(* IEC 61131-3 sources: courses/root/cat/cat-hw-boards/safety-plc/proj-safety-plc-emergency-stop-integration/structured-text, 4 files *)

(* ---- SafetyTypes.st ---- *)
TYPE E_SafetyState :
(
    STATE_SAFE := 0,               (* Безпечний робочий стан, силові виходи увімкнені *)
    STATE_ESTOP_ACTIVE := 1,        (* Натиснуто кнопку аварійної зупинки E-Stop (канали розімкнені) *)
    STATE_WAITING_FOR_RESET := 2,    (* Входи відновлено, очікується ручне підтвердження (Reset) *)
    STATE_DISCREPANCY_FAULT := 3,   (* Апаратна помилка: перевищено час розбіжності між каналами *)
    STATE_EDM_FAULT := 4            (* Апаратна помилка: несправність контактора або приварювання контактів *)
);
END_TYPE

TYPE E_EStopFault :
(
    ESTOP_FAULT_NONE := 0,                 (* Помилки відсутні *)
    ESTOP_FAULT_DISCREPANCY_TIMEOUT := 1,   (* Перевищення часу розбіжності спрацьовування каналів *)
    ESTOP_FAULT_EDM := 2,                   (* Несправність ланцюга зворотного зв'язку EDM *)
    ESTOP_FAULT_INVALID_RESET := 3          (* Некоректна послідовність скидання *)
);
END_TYPE

TYPE E_EdmFaultState :
(
    EDM_FAULT_NONE := 0,                (* Ланцюг зворотного зв'язку справний *)
    EDM_FAULT_CONTACT_WELDED := 1,      (* Приварювання контактів (NC не замкнувся при вимкненні) *)
    EDM_FAULT_CONTACT_STUCK_OPEN := 2,  (* Заклинювання реле (NC не розімкнувся при увімкненні) *)
    EDM_FAULT_TIMEOUT := 3              (* Таймаут підтвердження стану контакторів *)
);
END_TYPE

TYPE ST_EdmConfig :
STRUCT
    tFeedbackTimeout : TIME := T#250ms; (* Максимальний час очікування відповіді зворотного зв'язку *)
END_STRUCT
END_TYPE

TYPE ST_EStopConfig :
STRUCT
    tDiscrepancyTime : TIME := T#100ms; (* Допустима часова розбіжність між каналами E-Stop *)
    stEdmConfig      : ST_EdmConfig;    (* Конфігурація моніторингу зворотного зв'язку *)
END_STRUCT
END_TYPE

(* ---- FB_EDM_Monitor.st ---- *)
(*
    Функціональний блок: FB_EDM_Monitor
    Опис: Здійснює моніторинг зворотного зв'язку (External Device Monitoring) силових контакторів
          через їхні розмикальні (NC) допоміжні контакти. Забезпечує виявлення заклинювання
          або приварювання контактів за допомогою таймера контролю допустимої затримки перемикання.
*)
FUNCTION_BLOCK FB_EDM_Monitor
VAR_INPUT
    bControlOutput : BOOL;          (* Сигнал керування силових виходів (TRUE = увімкнено, FALSE = вимкнено) *)
    bFeedbackNC    : BOOL;          (* Сигнал з розмикальних (NC) допоміжних контактів контактора *)
    bReset         : BOOL;          (* Сигнал скидання помилки EDM *)
    stConfig       : ST_EdmConfig;  (* Конфігурація таймаутів моніторингу *)
END_VAR
VAR_OUTPUT
    bEdmOk         : BOOL := FALSE; (* Прапор норми: TRUE = ланцюг зворотного зв'язку у належному стані *)
    bError         : BOOL := FALSE; (* Прапор фіксації апаратної помилки контакторів *)
    eFaultState    : E_EdmFaultState := E_EdmFaultState.EDM_FAULT_NONE; (* Тип діагностованої помилки *)
END_VAR
VAR
    timerDelay     : TON;           (* Таймер затримки перемикання контактів *)
    bMismatch      : BOOL;          (* Прапор розбіжності між командою та зворотним зв'язком *)
END_VAR

(*
    Логіка моніторингу:
    У стабільному стані стан NC-контакту має бути протилежним команді керування:
    - Якщо bControlOutput = FALSE (контактор знеструмлено), NC-контакт має замкнутися (bFeedbackNC = TRUE).
    - Якщо bControlOutput = TRUE (контактор під напругою), NC-контакт має розімкнутися (bFeedbackNC = FALSE).
    Якщо bControlOutput = bFeedbackNC, виникає невідповідність (bMismatch = TRUE).
*)
bMismatch := (bControlOutput = bFeedbackNC);

(* Запуск таймера перевірки затримки спрацьовування *)
timerDelay(IN := bMismatch AND NOT bError, PT := stConfig.tFeedbackTimeout);

(* Фіксація помилки у разі перевищення таймауту *)
IF timerDelay.Q THEN
    bError := TRUE;
    IF NOT bControlOutput AND NOT bFeedbackNC THEN
        (* Вихід вимкнено, але NC-контакт не замкнувся -> приварювання силових контактів *)
        eFaultState := E_EdmFaultState.EDM_FAULT_CONTACT_WELDED;
    ELSIF bControlOutput AND bFeedbackNC THEN
        (* Вихід увімкнено, але NC-контакт не розімкнувся -> заклинювання у розімкненому стані *)
        eFaultState := E_EdmFaultState.EDM_FAULT_CONTACT_STUCK_OPEN;
    ELSE
        eFaultState := E_EdmFaultState.EDM_FAULT_TIMEOUT;
    END_IF;
END_IF;

(* Обробка процедури скидання помилки *)
IF bReset THEN
    (* Скидання дозволено лише якщо команду вимкнено і NC-контакт дійсно відновлено (замкнено) *)
    IF NOT bControlOutput AND bFeedbackNC THEN
        bError := FALSE;
        eFaultState := E_EdmFaultState.EDM_FAULT_NONE;
    END_IF;
END_IF;

(* Формування підсумкового прапорця стану EDM *)
bEdmOk := NOT bError AND NOT timerDelay.Q AND NOT bMismatch;

END_FUNCTION_BLOCK

(* ---- FB_EStop.st ---- *)
(*
    Функціональний блок: FB_EStop
    Опис: Реалізує функціонал безпеки двоканального аварійного зупину (E-Stop) з перевіркою
          часової розбіжності входів (Discrepancy Time), інтегрованим моніторингом зворотного
          зв'язку силових реле (EDM) та детермінованим автоматом станів.
*)
FUNCTION_BLOCK FB_EStop
VAR_INPUT
    bChannel1      : BOOL;          (* Перший канал кнопки E-Stop (F-DI 1, NC) *)
    bChannel2      : BOOL;          (* Другий канал кнопки E-Stop (F-DI 2, NC) *)
    bFeedbackNC    : BOOL;          (* Зворотний зв'язок NC-контактів силових реле *)
    bReset         : BOOL;          (* Сигнал кнопки ручного підтвердження/скидання (Reset) *)
    stConfig       : ST_EStopConfig;(* Параметри затримок та конфігурація EDM *)
END_VAR
VAR_OUTPUT
    bSafetyOutput  : BOOL := FALSE; (* Вихід дозволу роботи силових ланцюгів (F-DO) *)
    bReadyForReset : BOOL := FALSE; (* Сигнал індикації готовності до скидання (очікування Reset) *)
    bError         : BOOL := FALSE; (* Прапор виявлення апаратної помилки *)
    eState         : E_SafetyState := E_SafetyState.STATE_ESTOP_ACTIVE; (* Поточний стан безпеки *)
    eFault         : E_EStopFault  := E_EStopFault.ESTOP_FAULT_NONE;    (* Поточна фіксована помилка *)
END_VAR
VAR
    fbEdm          : FB_EDM_Monitor;(* Екземпляр блоку моніторингу контакторів *)
    timerDiscrepancy: TON;          (* Таймер контролю часової розбіжності входів *)
    rTrigReset     : R_TRIG;        (* Визначник наростаючого фронту для сигналу Reset *)
END_VAR

(* Виявлення фронту сигналу скидання (захист від постійно затиснутої кнопки Reset) *)
rTrigReset(CLK := bReset);

(* Виклик підсистеми EDM моніторингу *)
fbEdm(
    bControlOutput := bSafetyOutput,
    bFeedbackNC    := bFeedbackNC,
    bReset         := bReset,
    stConfig       := stConfig.stEdmConfig
);

(* Таймер контролю часової розбіжності між двома каналами кнопки аварійної зупинки *)
timerDiscrepancy(
    IN := (bChannel1 <> bChannel2) AND (eState <> E_SafetyState.STATE_DISCREPANCY_FAULT),
    PT := stConfig.tDiscrepancyTime
);

(* Фіксація помилки часової розбіжності при перевищенні таймауту *)
IF timerDiscrepancy.Q THEN
    eState := E_SafetyState.STATE_DISCREPANCY_FAULT;
    eFault := E_EStopFault.ESTOP_FAULT_DISCREPANCY_TIMEOUT;
END_IF;

(* Обробка виникнення аварії у ланцюзі EDM *)
IF fbEdm.bError AND (eState <> E_SafetyState.STATE_DISCREPANCY_FAULT) THEN
    eState := E_SafetyState.STATE_EDM_FAULT;
    eFault := E_EStopFault.ESTOP_FAULT_EDM;
END_IF;

(* Автомат станів безпеки *)
CASE eState OF
    E_SafetyState.STATE_SAFE:
        bSafetyOutput := TRUE;
        bReadyForReset := FALSE;
        bError := FALSE;

        (* Реагування на зміну стану каналів E-Stop *)
        IF NOT bChannel1 OR NOT bChannel2 THEN
            bSafetyOutput := FALSE;
            IF NOT bChannel1 AND NOT bChannel2 THEN
                eState := E_SafetyState.STATE_ESTOP_ACTIVE;
            END_IF;
        END_IF;

    E_SafetyState.STATE_ESTOP_ACTIVE:
        bSafetyOutput := FALSE;
        bReadyForReset := FALSE;
        bError := FALSE;

        (* Перехід у стан очікування скидання після відновлення обох каналів *)
        IF bChannel1 AND bChannel2 THEN
            eState := E_SafetyState.STATE_WAITING_FOR_RESET;
        END_IF;

    E_SafetyState.STATE_WAITING_FOR_RESET:
        bSafetyOutput := FALSE;
        bReadyForReset := TRUE;
        bError := FALSE;

        (* Перевірка повторного розмикання входів E-Stop *)
        IF NOT bChannel1 OR NOT bChannel2 THEN
            bReadyForReset := FALSE;
            IF NOT bChannel1 AND NOT bChannel2 THEN
                eState := E_SafetyState.STATE_ESTOP_ACTIVE;
            END_IF;
        (* Ручне скидання за допомогою фронту сигналу Reset *)
        ELSIF rTrigReset.Q THEN
            IF fbEdm.bEdmOk THEN
                eState := E_SafetyState.STATE_SAFE;
                eFault := E_EStopFault.ESTOP_FAULT_NONE;
            ELSE
                eState := E_SafetyState.STATE_EDM_FAULT;
                eFault := E_EStopFault.ESTOP_FAULT_EDM;
            END_IF;
        END_IF;

    E_SafetyState.STATE_DISCREPANCY_FAULT:
        bSafetyOutput := FALSE;
        bReadyForReset := FALSE;
        bError := TRUE;

        (* Квитування помилки розбіжності можливе лише після повного натискання кнопки E-Stop (обидва канали FALSE) *)
        IF NOT bChannel1 AND NOT bChannel2 THEN
            eState := E_SafetyState.STATE_ESTOP_ACTIVE;
        END_IF;

    E_SafetyState.STATE_EDM_FAULT:
        bSafetyOutput := FALSE;
        bReadyForReset := FALSE;
        bError := TRUE;

        (* Спроба відновлення роботи при натисканні Reset, якщо контактори справні *)
        IF rTrigReset.Q THEN
            IF NOT fbEdm.bError AND bChannel1 AND bChannel2 THEN
                eState := E_SafetyState.STATE_WAITING_FOR_RESET;
                eFault := E_EStopFault.ESTOP_FAULT_NONE;
            END_IF;
        END_IF;
END_CASE;

END_FUNCTION_BLOCK

(* ---- MAIN_Safety.st ---- *)
(*
    Програма: MAIN_Safety
    Опис: Головна циклічна програма (Safety PRG) для програмованого логічного контролера
          безпеки (Safety PLC). Здійснює опитування безпечних входів F-DI, викликає
          функціональний блок E-Stop та керує виходами безпеки F-DO і світлосигнальною арматурою.
*)
PROGRAM MAIN_Safety
VAR
    (* Фізичні / логічні входи безпеки (F-DI - Safe Digital Inputs) *)
    i_bEStop_Ch1     : BOOL := TRUE;  (* Вхід каналу 1 грибка аварійної зупинки *)
    i_bEStop_Ch2     : BOOL := TRUE;  (* Вхід каналу 2 грибка аварійної зупинки *)
    i_bContactor_NC  : BOOL := TRUE;  (* Зворотний зв'язок NC-контактів силових реле *)
    i_bResetButton   : BOOL := FALSE; (* Сигнал кнопки ручного підтвердження/скидання *)

    (* Фізичні / логічні виходи безпеки (F-DO - Safe Digital Outputs) *)
    q_bSafetyEnable  : BOOL := FALSE; (* Вихід дозволу живлення силових приводів *)
    q_bResetLamp     : BOOL := FALSE; (* Світловий індикатор кнопки Reset (очікування підтвердження) *)
    q_bFaultLamp     : BOOL := FALSE; (* Світловий індикатор аварії / несправності *)

    (* Екземпляр функціонального блоку логіки безпеки *)
    fbEStopLogic     : FB_EStop;

    (* Конфігурація параметрів затримок *)
    stSafetyConfig   : ST_EStopConfig;

    (* Прапор первинної ініціалізації *)
    bInitialised     : BOOL := FALSE;
END_VAR

(* Первинне встановлення параметрів у першому циклі *)
IF NOT bInitialised THEN
    stSafetyConfig.tDiscrepancyTime := T#100ms;
    stSafetyConfig.stEdmConfig.tFeedbackTimeout := T#250ms;
    bInitialised := TRUE;
END_IF;

(* Цикличне виконання логіки безпечного аварійного зупину *)
fbEStopLogic(
    bChannel1   := i_bEStop_Ch1,
    bChannel2   := i_bEStop_Ch2,
    bFeedbackNC := i_bContactor_NC,
    bReset      := i_bResetButton,
    stConfig    := stSafetyConfig
);

(* Запис результатів у виходи безпеки F-DO *)
q_bSafetyEnable := fbEStopLogic.bSafetyOutput;
q_bResetLamp    := fbEStopLogic.bReadyForReset;
q_bFaultLamp    := fbEStopLogic.bError;

END_PROGRAM
